Fanuc KAREL source: KO00020.KL

PROGRAM KO00020
%NOLOCKGROUP
VAR
  P1: XYZWPREXT
  P2: XYZWPREXT
  P3: XYZWPREXT
  OUT: JOINTPOS
BEGIN
  OUT = FRAME(P1, P2, P3)
END KO00020
